(* PLC project Controlador_PI, The Mathworks, Inc. Simulink PLC Coder 26.2 *)
(* stored: companyURL www.mathworks.com, creationDateTime 2026-10-27T10:24:52, productRelease (R2026b) *)

FUNCTION_BLOCK Controlador
  VAR_INPUT
    ssMethodType : SINT;
    In1 : LREAL;
    In2 : LREAL;
  END_VAR
  VAR_OUTPUT
    Out1 : LREAL;
  END_VAR
  VAR
    rtb_Sum : LREAL;
    c_DiscreteTimeIntegrator_DS : LREAL;
  END_VAR

            

CASE ssMethodType OF
    0: 
        (* SystemInitialize for Atomic SubSystem: '<Root>/Controlador' *)
        (* InitializeConditions for DiscreteIntegrator: '<S1>/Discrete-Time Integrator' *)
        c_DiscreteTimeIntegrator_DS := 0.0;
        (* End of SystemInitialize for SubSystem: '<Root>/Controlador' *)
    1: 
        (* Outputs for Atomic SubSystem: '<Root>/Controlador' *)
        (* Sum: '<S1>/Sum' *)
        rtb_Sum := In1 - In2;
        (* Outport: '<Root>/Out1' incorporates:
         *  DiscreteIntegrator: '<S1>/Discrete-Time Integrator'
         *  Gain: '<S1>/Ganho proporcional'
         *  Sum: '<S1>/Sum1' *)
        Out1 := (1.1 * rtb_Sum) + c_DiscreteTimeIntegrator_DS;
        (* Update for DiscreteIntegrator: '<S1>/Discrete-Time Integrator' incorporates:
         *  Gain: '<S1>/Ganho integral' *)
        c_DiscreteTimeIntegrator_DS := ((1.83 * rtb_Sum) * 0.1) + c_DiscreteTimeIntegrator_DS;
        (* End of Outputs for SubSystem: '<Root>/Controlador' *)
END_CASE;



          
END_FUNCTION_BLOCK
